(* CODESYS project beveling.project

Project tree, tasks and I/O mapping:
  Device : AM523-0808TN, Shenzhen Inovance Control Technology, version 3.5.11.50
      settings: PersistentStartAdddr = 0; PersistentStartEndAddr = 524287; Mode = 1
    application Application
      libraries: Standard, * (System); CmpEventMgr, 3.5.8.0 (System); Component Manager, 3.5.9.0 (System); CmpApp, 3.5.11.0 (System); CmpIecTask, 3.5.9.0 (System)
      task ETHERCAT1 (cyclic, interval 2000 µs, priority 0) calls ETHERCAT1.EtherCAT_Task, PLC_PRG
      task MainTask (cyclic, interval 4 ms, priority 1) calls nothing
      global variables GVL_Motion
      TaskEventPreStart
      program PLC_PRG [ST]
      DifferentialMonitor
    HardWare Configuration
    Resources List
    ConfigStorage
    Network Configuration
      LocalBus Config
      EtherCAT Config
    Device Diagnosis
    Serial : 串行接口, 汇川技术股份有限公司, version 00.00.00.10
      COM : Serial Port, Inovance, version 00.00.00.10
          settings: Device = AM523-0808TN; devGuid = 'e48f0cf2-85a4-455f-a8e7-135d3403221f'
    CAN : CAN总线, INOVANCE, version 00.00.00.10
    ETHERCAT1 : EtherCAT Master SoftMotion, 3S - Smart Software Solutions GmbH, version 3.5.11.10
        settings:  = 0; MasterCycleTime = 2000; NetworkName = 'eth1'; SelectNetworkByName = TRUE; DisableTaskGeneration = True; SlaveArrayName = ADR(_EC1_Node)
      InoSV660N : SV660_1Axis_00915, Inovance, order no. InoSV660N, version Revision=16#00010000
          settings: Number of Outputs = 6; Number of Inputs = 10; Number of Infos about Outputs = 6; Number of Infos about Inputs = 10; Configuration address of the slave = 1; Sync.Length = 18; Sync.Length = 32; FMMU.Length = 18; FMMU.Length = 32; DC sync0 cycletime = 2000; DC sync1 cycletime = 2000; Number of SDO = 10; Homing method.Index = 16#6098; Homing method.Subindex = 16#00; Homing method.Value = 1; Homing method.Size = 8; Homing method.AbortIfError = FALSE; Homing method.JumpToLine = FALSE; Homing method.Line = 0; Homing method.CompleteAccess = FALSE; Actual Position Calculation Method.Index = 16#60E6; Actual Position Calculation Method.Subindex = 16#00; Actual Position Calculation Method.Value = 0; Actual Position Calculation Method.Size = 8; Actual Position Calculation Method.AbortIfError = FALSE; Actual Position Calculation Method.JumpToLine = FALSE; Actual Position Calculation Method.Line = 0; Actual Position Calculation Method.CompleteAccess = FALSE; Speed during search for switch.Index = 16#6099; Speed during search for switch.Subindex = 16#01; Speed during search for switch.Value = 1398102; Speed during search for switch.Size = 32; Speed during search for switch.AbortIfError = FALSE; Speed during search for switch.JumpToLine = FALSE; Speed during search for switch.Line = 0; Speed during search for switch.CompleteAccess = FALSE; Homing acceleration.Index = 16#609A; Homing acceleration.Subindex = 16#00; Homing acceleration.Value = 139810133; Homing acceleration.Size = 32;
            Homing acceleration.AbortIfError = FALSE; Homing acceleration.JumpToLine = FALSE; Homing acceleration.Line = 0; Homing acceleration.CompleteAccess = FALSE; Speed during search for zero.Index = 16#6099; Speed during search for zero.Subindex = 16#02; Speed during search for zero.Value = 139810; Speed during search for zero.Size = 32; Speed during search for zero.AbortIfError = FALSE; Speed during search for zero.JumpToLine = FALSE; Speed during search for zero.Line = 0; Speed during search for zero.CompleteAccess = FALSE; Time of home searching.Index = 16#2005; Time of home searching.Subindex = 16#24; Time of home searching.Value = 50000; Time of home searching.Size = 16; Time of home searching.AbortIfError = FALSE; Time of home searching.JumpToLine = FALSE; Time of home searching.Line = 0; Time of home searching.CompleteAccess = FALSE; Positive torque limit value.Index = 16#60E0; Positive torque limit value.Subindex = 16#00; Positive torque limit value.Value = 3500; Positive torque limit value.Size = 16; Positive torque limit value.AbortIfError = FALSE; Positive torque limit value.JumpToLine = FALSE; Positive torque limit value.Line = 0; Positive torque limit value.CompleteAccess = FALSE; Negative torque limit value.Index = 16#60E1; Negative torque limit value.Subindex = 16#00; Negative torque limit value.Value = 3500; Negative torque limit value.Size = 16; Negative torque limit value.AbortIfError = FALSE; Negative torque limit value.JumpToLine = FALSE; Negative torque limit value.Line = 0; Negative torque limit value.CompleteAccess = FALSE; Max profile velocity.Index = 16#607F; Max profile velocity.Subindex = 16#00; Max profile velocity.Value = 83886080; Max profile velocity.Size = 32;
            Max profile velocity.AbortIfError = FALSE; Max profile velocity.JumpToLine = FALSE; Max profile velocity.Line = 0; Max profile velocity.CompleteAccess = FALSE; RxTxPdo.NumberofEntries = 6; RxTxPdo.Sm = 2; Controlword.Index = 16#6040; Controlword.SubIndex = 0; Controlword.Size = 16; Controlword.DependOnSlot = false; Controlword.DependOnSlotGroup = false; Target position.Index = 16#607A; Target position.SubIndex = 0; Target position.Size = 32; Target position.DependOnSlot = false; Target position.DependOnSlotGroup = false; Touch probe function.Index = 16#60B8; Touch probe function.SubIndex = 0; Touch probe function.Size = 16; Touch probe function.DependOnSlot = false; Touch probe function.DependOnSlotGroup = false; Physical outputs.Index = 16#60FE; Physical outputs.SubIndex = 1; Physical outputs.Size = 32; Physical outputs.DependOnSlot = false; Physical outputs.DependOnSlotGroup = false; Target velocity.Index = 16#60FF; Target velocity.SubIndex = 0; Target velocity.Size = 32; Target velocity.DependOnSlot = false; Target velocity.DependOnSlotGroup = false; Target torque.Index = 16#6071; Target torque.SubIndex = 0; Target torque.Size = 16; Target torque.DependOnSlot = false; Target torque.DependOnSlotGroup = false; RxTxPdo.Sm = -1; RxTxPdo.NumberofEntries = 10; RxTxPdo.Sm = 3; Error code.Index = 16#603F;
            Error code.SubIndex = 0; Error code.Size = 16; Error code.DependOnSlot = false; Error code.DependOnSlotGroup = false; Statusword.Index = 16#6041; Statusword.SubIndex = 0; Statusword.Size = 16; Statusword.DependOnSlot = false; Statusword.DependOnSlotGroup = false; Position actual value.Index = 16#6064; Position actual value.SubIndex = 0; Position actual value.Size = 32; Position actual value.DependOnSlot = false; Position actual value.DependOnSlotGroup = false; Torque actual value.Index = 16#6077; Torque actual value.SubIndex = 0; Torque actual value.Size = 16; Torque actual value.DependOnSlot = false; Torque actual value.DependOnSlotGroup = false; Following error actual value.Index = 16#60F4; Following error actual value.SubIndex = 0; Following error actual value.Size = 32; Following error actual value.DependOnSlot = false; Following error actual value.DependOnSlotGroup = false; Touch probe status.Index = 16#60B9; Touch probe status.SubIndex = 0; Touch probe status.Size = 16; Touch probe status.DependOnSlot = false; Touch probe status.DependOnSlotGroup = false; Touch probe pos1 pos value.Index = 16#60BA; Touch probe pos1 pos value.SubIndex = 0; Touch probe pos1 pos value.Size = 32; Touch probe pos1 pos value.DependOnSlot = false; Touch probe pos1 pos value.DependOnSlotGroup = false; Touch probe pos2 pos value.Index = 16#60BC; Touch probe pos2 pos value.SubIndex = 0; Touch probe pos2 pos value.Size = 32; Touch probe pos2 pos value.DependOnSlot = false; Touch probe pos2 pos value.DependOnSlotGroup = false; Digital inputs.Index = 16#60FD;
            Digital inputs.SubIndex = 0; Digital inputs.Size = 32; Digital inputs.DependOnSlot = false; Digital inputs.DependOnSlotGroup = false; Velocity actual value.Index = 16#606C; Velocity actual value.SubIndex = 0; Velocity actual value.Size = 32; Velocity actual value.DependOnSlot = false; Velocity actual value.DependOnSlotGroup = false; RxTxPdo.Sm = -1; Controlword.Name = 'Controlword'; Controlword.DataType = 'UINT'; Target position.Name = 'Target position'; Target position.DataType = 'DINT'; Touch probe function.Name = 'Touch probe function'; Touch probe function.DataType = 'UINT'; Physical outputs.Name = 'Physical outputs'; Physical outputs.DataType = 'UDINT'; Target velocity.Name = 'Target velocity'; Target velocity.DataType = 'DINT'; Target torque.Name = 'Target torque'; Target torque.DataType = 'INT'; Error code.Name = 'Error code'; Error code.DataType = 'UINT'; Statusword.Name = 'Statusword'; Statusword.DataType = 'UINT'; Position actual value.Name = 'Position actual value'; Position actual value.DataType = 'DINT'; Torque actual value.Name = 'Torque actual value'; Torque actual value.DataType = 'INT'; Following error actual value.Name = 'Following error actual value'; Following error actual value.DataType = 'DINT'; Touch probe status.Name = 'Touch probe status'; Touch probe status.DataType = 'UINT'; Touch probe pos1 pos value.Name = 'Touch probe pos1 pos value'; Touch probe pos1 pos value.DataType = 'DINT'; Touch probe pos2 pos value.Name = 'Touch probe pos2 pos value'; Touch probe pos2 pos value.DataType = 'DINT'; Digital inputs.Name = 'Digital inputs'; Digital inputs.DataType = 'UDINT';
            Velocity actual value.Name = 'Velocity actual value'; Velocity actual value.DataType = 'DINT'
          unmapped channels: Controlword, Target position, Touch probe function, Physical outputs, Target velocity, Target torque, Error code, Statusword, Position actual value, Torque actual value, Following error actual value, Touch probe status, Touch probe pos1 pos value, Touch probe pos2 pos value, Digital inputs, Velocity actual value
        Axis_1 : Axis, 3S - Smart Software Solutions GmbH, order no. 0, version 4.0.0.0
            settings: wDriveID = 0; dwRatioTechUnitsDenom = 4194304; iRatioTechUnitsNum = 5; HomingMode = 10; ZeroSignal = 0; StartDirction = 1; EndDirection = 1; PosLimitMode = 0; NegLimitMode = 0; HomingVelocity = 10; HomingApproachVelocity = 2; HomingAcceleration = 100; HomingDeceleration = 100; HomingJerk = 0; HomeMaskDistance = 0; HomePositionOffset = 0; HomePushTime = 0; HomeCompensation = 0; HomeTimeout = 0; HomeCompensationVelocity = 1000; 4000 = 1; 4001 = 0; 4003 = true; 4004 = 3; 4005 = 0; 4006 = 1.666667; 4007 = 166.666666; 4008 = 0.166667; 4009 = 50000; 4010 = 3500; 4011 = 3500; 4012 = 100.000000; ScalingIncs = 16#800000; 6005 = 10; AdrOffset_8010 = 4; BitOffset_8010 = 0; BitLength_8010 = 16; Address_8010 = '%QW2'; Type_8010 = 'UINT'; AddressPointer_8010 = ADR(%QW2);
              AdrOffset_8020 = 8; BitOffset_8020 = 0; BitLength_8020 = 32; Address_8020 = '%QD2'; Type_8020 = 'DINT'; AddressPointer_8020 = ADR(%QD2); AdrOffset_8030 = 20; BitOffset_8030 = 0; BitLength_8030 = 32; Address_8030 = '%QD5'; Type_8030 = 'DINT'; AddressPointer_8030 = ADR(%QD5); AdrOffset_8040 = 24; BitOffset_8040 = 0; BitLength_8040 = 16; Address_8040 = '%QW12'; Type_8040 = 'INT'; AddressPointer_8040 = ADR(%QW12); AdrOffset_8050 = 4294967295; BitOffset_8050 = 0; BitLength_8050 = 0; Address_8050 = ''; Type_8050 = ''; AddressPointer_8050 = 0; AdrOffset_8060 = 12; BitOffset_8060 = 0; BitLength_8060 = 16; Address_8060 = '%QW6'; Type_8060 = 'UINT'; AddressPointer_8060 = ADR(%QW6); AdrOffset_8070 = 4294967295; BitOffset_8070 = 0; BitLength_8070 = 0; Address_8070 = ''; Type_8070 = ''; AddressPointer_8070 = 0; AdrOffset_8080 = 4294967295; BitOffset_8080 = 0; BitLength_8080 = 0; Address_8080 = '';
              Type_8080 = ''; AddressPointer_8080 = 0; AdrOffset_8090 = 16; BitOffset_8090 = 0; BitLength_8090 = 32; Address_8090 = '%QD4'; Type_8090 = 'UDINT'; AddressPointer_8090 = ADR(%QD4); AdrOffset_8100 = 4294967295; BitOffset_8100 = 0; BitLength_8100 = 0; Address_8100 = ''; Type_8100 = ''; AddressPointer_8100 = 0; AdrOffset_8510 = 6; BitOffset_8510 = 0; BitLength_8510 = 16; Address_8510 = '%IW3'; Type_8510 = 'UINT'; AddressPointer_8510 = ADR(%IW3); AdrOffset_8520 = 8; BitOffset_8520 = 0; BitLength_8520 = 32; Address_8520 = '%ID2'; Type_8520 = 'DINT'; AddressPointer_8520 = ADR(%ID2); AdrOffset_8530 = 36; BitOffset_8530 = 0; BitLength_8530 = 32; Address_8530 = '%ID9'; Type_8530 = 'DINT'; AddressPointer_8530 = ADR(%ID9); AdrOffset_8540 = 12; BitOffset_8540 = 0; BitLength_8540 = 16; Address_8540 = '%IW6'; Type_8540 = 'INT'; AddressPointer_8540 = ADR(%IW6); AdrOffset_8550 = 4294967295; BitOffset_8550 = 0;
              BitLength_8550 = 0; Address_8550 = ''; Type_8550 = ''; AddressPointer_8550 = 0; AdrOffset_8560 = 32; BitOffset_8560 = 0; BitLength_8560 = 32; Address_8560 = '%ID8'; Type_8560 = 'UDINT'; AddressPointer_8560 = ADR(%ID8); AdrOffset_8570 = 20; BitOffset_8570 = 0; BitLength_8570 = 16; Address_8570 = '%IW10'; Type_8570 = 'UINT'; AddressPointer_8570 = ADR(%IW10); AdrOffset_8580 = 24; BitOffset_8580 = 0; BitLength_8580 = 32; Address_8580 = '%ID6'; Type_8580 = 'DINT'; AddressPointer_8580 = ADR(%ID6); AdrOffset_8590 = 4294967295; BitOffset_8590 = 0; BitLength_8590 = 0; Address_8590 = ''; Type_8590 = ''; AddressPointer_8590 = 0; AdrOffset_8600 = 28; BitOffset_8600 = 0; BitLength_8600 = 32; Address_8600 = '%ID7'; Type_8600 = 'DINT'; AddressPointer_8600 = ADR(%ID7); AdrOffset_8600 = 4294967295; BitOffset_8600 = 0; BitLength_8600 = 0; Address_8610 = ''; Type_8610 = ''; AddressPointer_8610 = 0;
              AdrOffset_8620 = 4; BitOffset_8620 = 0; BitLength_8620 = 16; Address_8620 = '%IW2'; Type_8620 = 'UINT'; AddressPointer_8620 = ADR(%IW2); IsValid = True; AxisNumber = 1; IsHostHoming = True; PulseSelectIndex = 4; SERVO_MAX_ID = 83886080
    EXP_A : 扩展卡, 汇川技术股份有限公司, version 00.00.00.10
    Local Bus
    MODBUS_TCP : ModbusTCP本地从站, inovance, version 00.00.00.10
    LocalHSIO : 本地高速IO, 汇川技术股份有限公司, version 2.0.0.0
        unmapped channels: DigitalInput, DigitalOutput
    HwConfiguratioinDevice : SystemConfig, Inovance, version 00.00.00.10
        settings: NetworkConfigArray.NetworkConfigArray.BusType = 10; NetworkConfigArray.NetworkConfigArray.RackSum = 1; NetworkConfigArray.NetworkConfigArray.HardwareConfigArray.HardwareConfigArray.RackNo = 1
    EXP_B : 扩展卡, 汇川技术股份有限公司, version 00.00.00.10
    SoftMotion General Axis Pool
*)

// Device/Application/GVL_Motion
VAR_GLOBAL
    (* ================= Commands (HMI / online write) ================= *)
    xEnable     : BOOL;              (* power on / off the servo axis *)
    xReset      : BOOL;              (* reset axis error *)
    xStop       : BOOL;              (* stop and lock the axis *)
    xJogFwd     : BOOL;              (* jog forward (level) *)
    xJogRev     : BOOL;              (* jog reverse (level) *)
    xMoveRel    : BOOL;              (* relative move command (level) *)
    xMoveAbs    : BOOL;              (* absolute move command (level) *)
    xStartCycle : BOOL;              (* start auto fwd/back cycle (rising edge) *)

    rRelDist    : LREAL := 100.0;    (* relative move distance [mm] *)
    rTargetPos  : LREAL := 0.0;      (* absolute target position [mm] *)

    (* ================= Motion parameters ================= *)
    rJogVel     : LREAL := 10.0;     (* jog velocity [mm/s] *)
    rVel        : LREAL := 30.0;     (* positioning velocity [mm/s] *)
    rAcc        : LREAL := 200.0;    (* acceleration [mm/s2] *)
    rDec        : LREAL := 200.0;    (* deceleration [mm/s2] *)
    rStroke     : LREAL := 100.0;    (* auto cycle stroke (one way) [mm] *)
    tDwell      : TIME  := T#1S;     (* dwell time at cycle ends *)

    (* ================= Status ================= *)
    xPowered    : BOOL;              (* MC_Power.Status : servo enabled *)
    xAxisReady  : BOOL;              (* axis in StandStill -> motion allowed *)
    xBusy       : BOOL;              (* any motion active *)
    xDisabled   : BOOL;              (* axis state = Disabled *)
    xStandStill : BOOL;              (* axis state = StandStill *)
    xStopping   : BOOL;              (* axis state = Stopping *)
    xErrorStop  : BOOL;              (* axis state = ErrorStop *)
    xAxisError  : BOOL;              (* axis reports an error *)
    iAxisErrorID: DWORD;             (* axis error code *)
    rActPos     : LREAL;             (* actual position [mm] *)
    iState      : INT;               (* auto cycle step number *)
END_VAR

// Device/Application/PLC_PRG
PROGRAM PLC_PRG
VAR
    (* ---- SoftMotion function block instances ---- *)
    fbPower    : MC_Power;            (* enable / disable the axis *)
    fbReset    : MC_Reset;            (* reset axis error *)
    fbStop     : MC_Stop;             (* stop and lock the axis *)
    fbJog      : MC_Jog;              (* jog *)
    fbMoveRel  : MC_MoveRelative;     (* single relative move *)
    fbMoveAbs  : MC_MoveAbsolute;     (* single absolute move *)
    fbCycle    : MC_MoveRelative;     (* auto cycle move *)
    fbReadPos  : MC_ReadActualPosition; (* position feedback *)
    fbReadStat : MC_ReadStatus;       (* axis state machine *)
    fbReadErr  : MC_ReadAxisError;    (* axis error code *)

    (* ---- edge detection ---- *)
    rtCycle    : R_TRIG;              (* auto cycle trigger *)

    (* ---- auto cycle ---- *)
    fbCycleExec: BOOL;                (* Execute for fbCycle *)
    rCycleDist : LREAL;               (* current segment distance *)
    iCycle     : INT := 0;            (* auto cycle step *)
    tonDwell   : TON;                 (* dwell at cycle ends *)

    (* ---- diagnostics ---- *)
    eLastErr   : SMC_ERROR;           (* latched last motion block error *)
	xDoReset: BOOL;
	xStopRun: BOOL;
	rRunDec: LREAL;
	xStartRun: BOOL;
	iStep: INT;
	fbMoveVel: MC_MoveVelocity;
	Axis: INT;
	Execute: BOOL;
	rRunVel: LREAL;
	rRunAcc: LREAL;
	Velocity: INT;
	Acceleration: INT;
	Deceleration: INT;
	Direction: INT;
	InVelocity: INT;
	xMoveExec: BOOL;
END_VAR

(* Single low-speed 20 mm out-and-back test cycle.
   Start only on a rising edge of GVL_Motion.xStartCycle.
   Travel is capped at 20 mm per leg and 10 mm/s. *)
rtCycle(CLK := GVL_Motion.xStartCycle);

fbPower(Axis         := Axis_1,
        Enable       := GVL_Motion.xEnable,
        bRegulatorOn := TRUE,
        bDriveStart  := TRUE);

fbReset(Axis := Axis_1, Execute := GVL_Motion.xReset);

IF GVL_Motion.xStop THEN
    xStopRun   := TRUE;
    fbCycleExec := FALSE;
    iCycle      := 0;
END_IF

IF fbPower.Error OR fbCycle.Error OR fbReset.Error OR fbStop.Error THEN
    iCycle      := 99;
    fbCycleExec := FALSE;
    xStopRun    := TRUE;
END_IF

fbStop(Axis         := Axis_1,
       Execute      := xStopRun,
       Deceleration := MIN(MAX(GVL_Motion.rDec, 10.0), 200.0));

IF xStopRun AND fbStop.Done THEN
    xStopRun := FALSE;
END_IF

tonDwell(IN := (iCycle = 20) OR (iCycle = 40),
         PT := GVL_Motion.tDwell);

CASE iCycle OF
    0:  (* Idle; one rising edge starts one round trip. *)
        fbCycleExec := FALSE;
        IF rtCycle.Q
           AND GVL_Motion.xEnable
           AND fbPower.Status
           AND NOT GVL_Motion.xAxisError
           AND NOT xStopRun
           AND (ABS(GVL_Motion.rStroke) > 0.0) THEN
            rCycleDist := MIN(ABS(GVL_Motion.rStroke), 20.0);
            fbCycleExec := TRUE;
            iCycle := 10;
        END_IF

    10: (* Forward leg. *)
        IF fbCycle.Done THEN
            fbCycleExec := FALSE;
            iCycle := 20;
        ELSIF fbCycle.Error THEN
            fbCycleExec := FALSE;
            iCycle := 99;
            xStopRun := TRUE;
        END_IF

    20: (* Dwell before return leg. *)
        IF tonDwell.Q AND NOT xStopRun THEN
            rCycleDist := -MIN(ABS(GVL_Motion.rStroke), 20.0);
            fbCycleExec := TRUE;
            iCycle := 30;
        END_IF

    30: (* Return leg. *)
        IF fbCycle.Done THEN
            fbCycleExec := FALSE;
            iCycle := 40;
        ELSIF fbCycle.Error THEN
            fbCycleExec := FALSE;
            iCycle := 99;
            xStopRun := TRUE;
        END_IF

    40: (* Dwell after returning to the start position, then finish. *)
        IF tonDwell.Q THEN
            iCycle := 0;
        END_IF

    99: (* Error latch; require a successful reset and completed stop. *)
        fbCycleExec := FALSE;
        IF GVL_Motion.xReset AND fbReset.Done AND NOT xStopRun THEN
            iCycle := 0;
        END_IF

ELSE
    iCycle := 99;
    fbCycleExec := FALSE;
    xStopRun := TRUE;
END_CASE

fbCycle(Axis         := Axis_1,
        Execute      := fbCycleExec AND NOT xStopRun,
        Distance     := rCycleDist,
        Velocity     := MIN(MAX(GVL_Motion.rVel, 1.0), 10.0),
        Acceleration := MIN(MAX(GVL_Motion.rAcc, 10.0), 200.0),
        Deceleration := MIN(MAX(GVL_Motion.rDec, 10.0), 200.0));

fbReadPos(Axis := Axis_1, Enable := TRUE);

GVL_Motion.xPowered    := fbPower.Status;
GVL_Motion.xBusy       := fbCycle.Busy OR fbStop.Busy;
GVL_Motion.xDisabled   := NOT fbPower.Status;
GVL_Motion.xStopping   := fbStop.Busy;
GVL_Motion.xStandStill := fbPower.Status AND NOT GVL_Motion.xBusy;
GVL_Motion.xAxisReady  := GVL_Motion.xStandStill AND NOT GVL_Motion.xAxisError;
GVL_Motion.xAxisError  := fbPower.Error OR fbCycle.Error OR fbReset.Error OR fbStop.Error;
GVL_Motion.xErrorStop  := GVL_Motion.xAxisError;
GVL_Motion.iState      := iCycle;
GVL_Motion.rActPos     := fbReadPos.Position;

END_PROGRAM
